(* IEC 61131-3 sources: ZPLC/packages/zplc-ide/projects/two_hand/src, 1 file *)

(* ---- TwoHand.st ---- *)
PROGRAM TwoHand
VAR_INPUT LeftHand AT %I0.0 : BOOL; RightHand AT %I0.1 : BOOL; GuardClosed AT %I0.2 : BOOL; END_VAR
VAR_OUTPUT PressEnable AT %Q0.0 : BOOL; GuardLamp AT %Q0.1 : BOOL; OneHandWarning AT %Q0.2 : BOOL; END_VAR
PressEnable := LeftHand AND RightHand AND GuardClosed; GuardLamp := NOT GuardClosed; OneHandWarning := LeftHand XOR RightHand;
END_PROGRAM
